(* IEC 61131-3 sources: plc-iiot-stack/tests/POUs/FB_IiotFunctions_Test, 4 files *)

(* ---- AlarmStateFromWords.method.decl.st ---- *)
// Состояние тревоги по словам: OOS, подавлена, отложена, активна/неквитирована, вернулась, норма.
METHOD PRIVATE AlarmStateFromWords
VAR
    stWords : ST_IiotAlarmWords;
END_VAR

(* ---- NonFiniteTransitionsAreChanges.method.decl.st ---- *)
// Переход между числом и NaN/бесконечностью — изменение; два неконечных — нет.
METHOD PRIVATE NonFiniteTransitionsAreChanges
VAR
    lwNan : LWORD := 16#7FF8000000000000;
    lwInf : LWORD := 16#7FF0000000000000;
    pBits : POINTER TO LREAL;
    lrNan : LREAL;
    lrInf : LREAL;
END_VAR

(* ---- NowIsMonotonic.method.decl.st ---- *)
// Монотонное время: время с запуска больше нуля, повторный вызов не возвращает меньшее значение.
METHOD PRIVATE NowIsMonotonic
VAR
    ltFirst : LTIME;
    ltSecond : LTIME;
END_VAR

(* ---- ZeroNegativeOrNanDeadbandMeansAnyChange.method.decl.st ---- *)
// Зона <= 0 или не число — любое изменение.
METHOD PRIVATE ZeroNegativeOrNanDeadbandMeansAnyChange
VAR
    dwNan : DWORD := 16#7FC00000;
    pBitsR : POINTER TO REAL;
    rNan : REAL;
END_VAR
